// TIA Portal V20 export
DATA_BLOCK "T7_Resultado"   // DB44901
{ S7_Optimized_Access := 'TRUE' }
AUTHOR : IA
FAMILY : PRUEBA
VERSION : 0.1
// Tanda 3: un Bool por prueba
// stored: AutoNumber false
   VAR
      L_JMP : Bool;   // JMP + LABEL (JumpCoil, Label)
      L_JMPN : Bool;   // JMPN (I_JumpCoil)
      L_JMP_LIST : Bool;   // JMP_LIST (JumpList), K = 1
      L_SWITCH : Bool;   // SWITCH (Switch), K = 5 → caso 1
      L_RE_TRIGR : Bool;   // RE_TRIGR
      L_GET_ERROR : Bool;   // GET_ERROR (GetError) y GET_ERR_ID (GetErrorID) sin error
      L_WAIT : Bool;   // WAIT
      L_VariantGet : Bool;   // VariantGet (Variant → Int)
      L_VariantPut : Bool;   // VariantPut (Int → Variant)
      L_ArrayDB : Bool;   // WriteToArrayDB + ReadFromArrayDB
      L_ATTR_DB : Bool;   // ATTR_DB sobre T7_Std (longitud > 0)
      L_AIRT : Bool;   // DIS_AIRT + EN_AIRT
      L_SRT_DINT : Bool;   // SRT_DINT + QRY_DINT: el OB20 se ha ejecutado
      L_QRY_CINT : Bool;   // QRY_CINT y el OB30 se ejecuta
      L_Program_Alarm : Bool;   // Program_Alarm sin error
      L_RTM : Bool;   // RTM modo 0 (leer)
      S_PEEK_POKE : Bool;   // [SCL] POKE + PEEK en un DB de acceso estándar
      S_BIG_LITTLE : Bool;   // [SCL] WRITE_BIG/READ_BIG y WRITE_LITTLE/READ_LITTLE
      S_ArrayDB : Bool;   // [SCL] WriteToArrayDB / ReadFromArrayDB
      S_Variant : Bool;   // [SCL] VariantGet / VariantPut, TypeOf
      Vida : DInt;   // Sube cada ciclo
      OK : Int;   // Correctas
      Total : Int := 20;   // Pruebas
      Todo_OK : Bool;   // Todas correctas
   END_VAR
BEGIN
END_DATA_BLOCK
